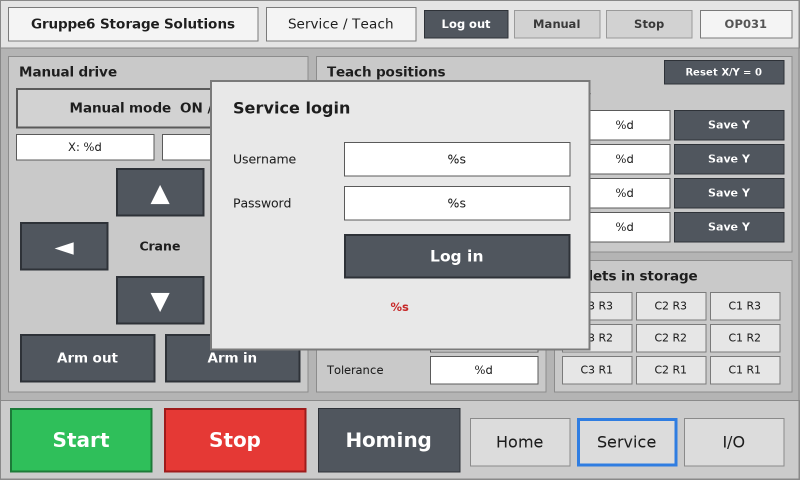
VISUALIZATION Service  // 800x480
    Rectangle (0,0 800x480)
    Rectangle (0,0 800x48)
    Rectangle (8,7 250x34), "Gruppe6 Storage Solutions"
    Rectangle (266,7 150x34), "Service / Teach"
    Rectangle (514,10 86x28), "Manual", colour toggle: MAIN.isManualMode
    Rectangle (606,10 86x28), "Stop", colour toggle: MAIN.isStop
    Rectangle (700,10 92x28), "OP031"
    Rectangle (0,400 800x80)
    RoundedRectangle (10,408 142x64), "Start"
        OnMouseUp: execute { MAIN.isStop := FALSE; }
    RoundedRectangle (164,408 142x64), "Stop"
        OnMouseUp: execute { MAIN.isStop := TRUE; }
    Rectangle (470,418 100x48), "Home"
        OnMouseUp: execute {
            MAIN.logoutRequest := TRUE;   // leaving the service page logs out
        }
        OnMouseUp: change screen: Start
    Rectangle (577,418 100x48), "Service"
        OnMouseUp: change screen: Service
    RoundedRectangle (424,10 84x28), "Log out", invisible if: MAIN.isServiceLocked, input disabled if: MAIN.isServiceLocked
        OnMouseUp: execute { MAIN.logoutRequest := TRUE; }
    Rectangle (8,56 300x336), invisible if: MAIN.isServiceLocked
    Rectangle (16,60 284x24), "Manual drive", invisible if: MAIN.isServiceLocked
    RoundedRectangle (16,88 284x40), "Manual mode ON / OFF", colour toggle: MAIN.isManualMode, invisible if: MAIN.isServiceLocked, input disabled if: MAIN.isServiceLocked
        toggle MAIN.isManualMode
    Rectangle (16,134 138x26), "X: %d", text variable: MAIN.currentPosX, invisible if: MAIN.isServiceLocked
    Rectangle (162,134 138x26), "Y: %d", text variable: MAIN.currentPosY, invisible if: MAIN.isServiceLocked
    RoundedRectangle (116,168 88x48), "▲", invisible if: MAIN.isServiceLocked, input disabled if: MAIN.isServiceLocked
        tap MAIN.jogUp
    RoundedRectangle (20,222 88x48), "◄", invisible if: MAIN.isServiceLocked, input disabled if: MAIN.isServiceLocked
        tap MAIN.jogToRack
    Rectangle (116,222 88x48), "Crane", invisible if: MAIN.isServiceLocked
    RoundedRectangle (212,222 88x48), "►", invisible if: MAIN.isServiceLocked, input disabled if: MAIN.isServiceLocked
        tap MAIN.jogToConveyor
    RoundedRectangle (116,276 88x48), "▼", invisible if: MAIN.isServiceLocked, input disabled if: MAIN.isServiceLocked
        tap MAIN.jogDown
    RoundedRectangle (20,334 135x48), "Arm out", invisible if: MAIN.isServiceLocked, input disabled if: MAIN.isServiceLocked
        tap MAIN.jogArmOut
    RoundedRectangle (165,334 135x48), "Arm in", invisible if: MAIN.isServiceLocked, input disabled if: MAIN.isServiceLocked
        tap MAIN.jogArmIn
    Rectangle (316,56 476x196), invisible if: MAIN.isServiceLocked
    Rectangle (324,60 300x24), "Teach positions", invisible if: MAIN.isServiceLocked
    RoundedRectangle (664,60 120x24), "Reset X/Y = 0", invisible if: MAIN.isServiceLocked, input disabled if: MAIN.isServiceLocked
        OnMouseUp: execute {
            // Set the position to zero (use it when the crane stands at the reference switches)
            MAIN.currentPosX := 0;
            MAIN.currentPosY := 0;
        }
    RoundedRectangle (318,408 142x64), "Homing", colour toggle: MAIN.isHoming, invisible if: MAIN.isServiceLocked, input disabled if: MAIN.isServiceLocked
        OnMouseUp: execute {
            MAIN.homeRequest := TRUE;   // start homing: arm in, crane to B1 and B4, position := 0
        }
    Rectangle (324,88 80x20), "Slot", invisible if: MAIN.isServiceLocked
    Rectangle (408,88 90x20), "X", invisible if: MAIN.isServiceLocked
    Rectangle (580,88 90x20), "Y", invisible if: MAIN.isServiceLocked
    Rectangle (324,110 80x30), "Conv. (0)", invisible if: MAIN.isServiceLocked
    Rectangle (408,110 90x30), "%d", text variable: MAIN.xPosition[0], invisible if: MAIN.isServiceLocked, input disabled if: MAIN.isServiceLocked
        OnMouseUp: write the text variable via Default
    RoundedRectangle (502,110 74x30), "Save X", invisible if: MAIN.isServiceLocked, input disabled if: MAIN.isServiceLocked
        OnMouseUp: execute {
            MAIN.xPosition[0] := MAIN.currentPosX;   // teach X
        }
    Rectangle (580,110 90x30), "%d", text variable: MAIN.yPosition[0], invisible if: MAIN.isServiceLocked, input disabled if: MAIN.isServiceLocked
        OnMouseUp: write the text variable via Default
    RoundedRectangle (674,110 110x30), "Save Y", invisible if: MAIN.isServiceLocked, input disabled if: MAIN.isServiceLocked
        OnMouseUp: execute {
            MAIN.yPosition[0] := MAIN.currentPosY;   // teach Y
        }
    Rectangle (324,144 80x30), "C1 / R1", invisible if: MAIN.isServiceLocked
    Rectangle (408,144 90x30), "%d", text variable: MAIN.xPosition[1], invisible if: MAIN.isServiceLocked, input disabled if: MAIN.isServiceLocked
        OnMouseUp: write the text variable via Default
    RoundedRectangle (502,144 74x30), "Save X", invisible if: MAIN.isServiceLocked, input disabled if: MAIN.isServiceLocked
        OnMouseUp: execute {
            MAIN.xPosition[1] := MAIN.currentPosX;   // teach X
        }
    Rectangle (580,144 90x30), "%d", text variable: MAIN.yPosition[1], invisible if: MAIN.isServiceLocked, input disabled if: MAIN.isServiceLocked
        OnMouseUp: write the text variable via Default
    RoundedRectangle (674,144 110x30), "Save Y", invisible if: MAIN.isServiceLocked, input disabled if: MAIN.isServiceLocked
        OnMouseUp: execute {
            MAIN.yPosition[1] := MAIN.currentPosY;   // teach Y
        }
    Rectangle (324,178 80x30), "C2 / R2", invisible if: MAIN.isServiceLocked
    Rectangle (408,178 90x30), "%d", text variable: MAIN.xPosition[2], invisible if: MAIN.isServiceLocked, input disabled if: MAIN.isServiceLocked
        OnMouseUp: write the text variable via Default
    RoundedRectangle (502,178 74x30), "Save X", invisible if: MAIN.isServiceLocked, input disabled if: MAIN.isServiceLocked
        OnMouseUp: execute {
            MAIN.xPosition[2] := MAIN.currentPosX;   // teach X
        }
    Rectangle (580,178 90x30), "%d", text variable: MAIN.yPosition[2], invisible if: MAIN.isServiceLocked, input disabled if: MAIN.isServiceLocked
        OnMouseUp: write the text variable via Default
    RoundedRectangle (674,178 110x30), "Save Y", invisible if: MAIN.isServiceLocked, input disabled if: MAIN.isServiceLocked
        OnMouseUp: execute {
            MAIN.yPosition[2] := MAIN.currentPosY;   // teach Y
        }
    Rectangle (324,212 80x30), "C3 / R3", invisible if: MAIN.isServiceLocked
    Rectangle (408,212 90x30), "%d", text variable: MAIN.xPosition[3], invisible if: MAIN.isServiceLocked, input disabled if: MAIN.isServiceLocked
        OnMouseUp: write the text variable via Default
    RoundedRectangle (502,212 74x30), "Save X", invisible if: MAIN.isServiceLocked, input disabled if: MAIN.isServiceLocked
        OnMouseUp: execute {
            MAIN.xPosition[3] := MAIN.currentPosX;   // teach X
        }
    Rectangle (580,212 90x30), "%d", text variable: MAIN.yPosition[3], invisible if: MAIN.isServiceLocked, input disabled if: MAIN.isServiceLocked
        OnMouseUp: write the text variable via Default
    RoundedRectangle (674,212 110x30), "Save Y", invisible if: MAIN.isServiceLocked, input disabled if: MAIN.isServiceLocked
        OnMouseUp: execute {
            MAIN.yPosition[3] := MAIN.currentPosY;   // teach Y
        }
    Rectangle (316,260 230x132), invisible if: MAIN.isServiceLocked
    Rectangle (324,264 210x24), "Parameters", invisible if: MAIN.isServiceLocked
    Rectangle (324,292 100x28), "Lift", invisible if: MAIN.isServiceLocked
    Rectangle (430,292 108x28), "%d", text variable: MAIN.liftOffset, invisible if: MAIN.isServiceLocked, input disabled if: MAIN.isServiceLocked
        OnMouseUp: write the text variable via Default
    Rectangle (324,324 100x28), "Lower", invisible if: MAIN.isServiceLocked
    Rectangle (430,324 108x28), "%d", text variable: MAIN.lowerOffset, invisible if: MAIN.isServiceLocked, input disabled if: MAIN.isServiceLocked
        OnMouseUp: write the text variable via Default
    Rectangle (324,356 100x28), "Tolerance", invisible if: MAIN.isServiceLocked
    Rectangle (430,356 108x28), "%d", text variable: MAIN.tolerance, invisible if: MAIN.isServiceLocked, input disabled if: MAIN.isServiceLocked
        OnMouseUp: write the text variable via Default
    Rectangle (554,260 238x132), invisible if: MAIN.isServiceLocked
    Rectangle (562,264 222x24), "Pallets in storage", invisible if: MAIN.isServiceLocked
    Rectangle (562,292 70x28), "C3 R3", colour toggle: MAIN.slotOccupied[3,3], invisible if: MAIN.isServiceLocked, input disabled if: MAIN.isServiceLocked
        toggle MAIN.slotOccupied[3,3]
    Rectangle (636,292 70x28), "C2 R3", colour toggle: MAIN.slotOccupied[2,3], invisible if: MAIN.isServiceLocked, input disabled if: MAIN.isServiceLocked
        toggle MAIN.slotOccupied[2,3]
    Rectangle (710,292 70x28), "C1 R3", colour toggle: MAIN.slotOccupied[1,3], invisible if: MAIN.isServiceLocked, input disabled if: MAIN.isServiceLocked
        toggle MAIN.slotOccupied[1,3]
    Rectangle (562,324 70x28), "C3 R2", colour toggle: MAIN.slotOccupied[3,2], invisible if: MAIN.isServiceLocked, input disabled if: MAIN.isServiceLocked
        toggle MAIN.slotOccupied[3,2]
    Rectangle (636,324 70x28), "C2 R2", colour toggle: MAIN.slotOccupied[2,2], invisible if: MAIN.isServiceLocked, input disabled if: MAIN.isServiceLocked
        toggle MAIN.slotOccupied[2,2]
    Rectangle (710,324 70x28), "C1 R2", colour toggle: MAIN.slotOccupied[1,2], invisible if: MAIN.isServiceLocked, input disabled if: MAIN.isServiceLocked
        toggle MAIN.slotOccupied[1,2]
    Rectangle (562,356 70x28), "C3 R1", colour toggle: MAIN.slotOccupied[3,1], invisible if: MAIN.isServiceLocked, input disabled if: MAIN.isServiceLocked
        toggle MAIN.slotOccupied[3,1]
    Rectangle (636,356 70x28), "C2 R1", colour toggle: MAIN.slotOccupied[2,1], invisible if: MAIN.isServiceLocked, input disabled if: MAIN.isServiceLocked
        toggle MAIN.slotOccupied[2,1]
    Rectangle (710,356 70x28), "C1 R1", colour toggle: MAIN.slotOccupied[1,1], invisible if: MAIN.isServiceLocked, input disabled if: MAIN.isServiceLocked
        toggle MAIN.slotOccupied[1,1]
    RoundedRectangle (210,80 380x270), invisible if: MAIN.isServiceUnlocked
    Rectangle (230,92 340x32), "Service login", invisible if: MAIN.isServiceUnlocked
    Rectangle (230,142 110x34), "Username", invisible if: MAIN.isServiceUnlocked
    Rectangle (344,142 226x34), "%s", text variable: MAIN.loginUser, invisible if: MAIN.isServiceUnlocked, input disabled if: MAIN.isServiceUnlocked
        OnMouseUp: write the text variable via Default, title 'Username'
    Rectangle (230,186 110x34), "Password", invisible if: MAIN.isServiceUnlocked
    Rectangle (344,186 226x34), "%s", text variable: MAIN.loginPasswordStars, invisible if: MAIN.isServiceUnlocked, input disabled if: MAIN.isServiceUnlocked
        OnMouseUp: write MAIN.loginPassword via Default, title 'Password', password
    RoundedRectangle (344,234 226x44), "Log in", invisible if: MAIN.isServiceUnlocked, input disabled if: MAIN.isServiceUnlocked
        OnMouseUp: execute { MAIN.loginRequest := TRUE; }
    Rectangle (230,292 340x30), "%s", text variable: MAIN.loginMessage, invisible if: MAIN.isServiceUnlocked
    Rectangle (684,418 100x48), "I/O", invisible if: MAIN.isServiceLocked, input disabled if: MAIN.isServiceLocked
        OnMouseUp: change screen: IO
END_VISUALIZATION

(* stored: Version 1.1.0.1, ProductVersion 3.1.4024.12
   Visu Service: Id {9470ee7a-673c-407b-8946-0c1fe32a4224} *)
